# EPICS IOC start-up script: examples/test/PSI/epp1008.iocsh
#- mXsXXX naming
require ecmccfg, "NAMING=mXsXXX"

#- add slaves
${SCRIPTEXEC} ${ecmccfg_DIR}addSlave.cmd, "HW_DESC=EPP1008, SLAVE_ID=2"
